(* IEC 61131-3 sources: Gen-AI/final/Gen-AI_v1.0_submission/A2_框架源码/agent/logs/full34_fixture/E3_P07_1_42/tools/candidate_1/fixture_compile, 1 file *)

(* ---- source.st ---- *)
TYPE ST_Pump :
STRUCT
    priority : INT;
    selection : BOOL;
    RunComd : BOOL;
END_STRUCT
END_TYPE
FUNCTION_BLOCK FB_P07
VAR_INPUT
    mode : BOOL;
    start : BOOL;
    stop : BOOL;
END_VAR
VAR_IN_OUT
    pumpGroup : ARRAY[1..5] OF ST_Pump;
END_VAR
(* Add a VAR block for internal state/timers before the implementation, if needed. *)
(* SKELETON ONLY: replace this RETURN with scan logic and required initial state. *)
RETURN;
END_FUNCTION_BLOCK

(* FIXTURE_COMPILE_FAIL *)
